(* IEC 61131-3 sources: codesys/project-view/Device/Plc Logic/Application/本机-3-机械臂-本体, 4 files *)

(* ---- Robot_STATE.st ---- *)
{attribute 'qualified_only'}
{attribute 'strict'}
(*A区三轴模组状态机*)
TYPE Robot_STATE :
(
	STOP := 0,						//停止
	INIT,						//初始化
	MANNUAL,					//手动模式
	AUTO,						//自动模式
	RobotAct,					//自动运行中
	MannualRun					//手动运行中
);
END_TYPE

(* ---- ST_ROBOT_MODULE.st ---- *)
TYPE ST_ROBOT_MODULE :	//机械臂模块
STRUCT
	bConnect					:BOOL;
	bConnected					:BOOL;
	bTcpError					:BOOL;

	//写
	x_iGrpEnable				:BOOL;			//上使能
	x_iGrpDisable				:BOOL;			//去使能
	x_iGrpReset					:BOOL;			//复位
	x_iStartScript				:BOOL;			//开始脚本
	x_iPauseScript				:BOOL;			//暂停脚本
	x_iContinueScript			:BOOL;			//继续脚本
	x_iStopScript				:BOOL;			//停止脚本
	x_iManualMode				:BOOL;			//手动模式
	x_iAutoMode					:BOOL;			//自动模式

	//读
	x_oStateRunning				:BOOL;			//状态-运行中
	x_oStateStopping			:BOOL;			//状态-停止中
	x_oStatePausing				:BOOL;			//状态-暂停中
	x_oStateFree				:BOOL;			//状态-空闲中
	x_oStateElectrify			:BOOL;			//状态-上电
	x_oStatePower				:BOOL;			//状态-使能中
	x_oStateErr					:BOOL;			//状态-报警
	x_oCollide					:BOOL;			//状态-碰撞

	//写
	wExecute_Init    			:WORD := 1;		//-- PLC请求初始化 (0/1)
	wExecute_Act     			:word;		//-- PLC请求执行动作 (0=无, 1=下料, 2=上料)
	wOrderNumCur     			:word;		//-- PLC指定工作站点 (1,2...)
	wRackTpye        			:word;		//-- PLC指定盘架类型
	wDeviceRackPosNum			:word;		//-- PLC指定设备取放编号
	wChassisRackPosNum			:WORD;		//-- PLC指定小车底盘位置编号
	xExcuteSetVal				:BOOL;		//搬运参数写入
	xExcuteInit					:BOOL;		//机械臂初始化
	xExcuteAct					:BOOL;		//执行机械臂搬运动作

	//读
	rGlobInitStatus				:WORD;			//初始化状态反馈		--4是初始化完成
	rOrderNumCur				:WORD;			//工作站点参数反馈
	rRackTpye					:WORD;			//盘架类型参数反馈
	rDeviceRackPosNum			:WORD;			//设备位置参数反馈
	rChassisRackPosNum			:WORD;			//小车位置参数反馈
	rAct_Status					:WORD;			//机械臂动作状态 (0=未执行,1=执行中,2=完成,3=失败)
	rExecute_Act				:WORD;			//当前执行动作反馈 (0=无, 1=下料, 2=上料)
	RobotBusy					:WORD;			//机械臂忙标志 (0=空闲, 1=忙碌)

	G_FailCode					:WORD;			//失败代码 (0=无错误, 1=RTU连接失败, 2=电爪初始化失败, 3=电爪打开失败, 4=电爪夹紧失败, 5=拍照失败)
	G_FailWorkstationrk			:WORD;			//失败时的工作站点编号
	G_FailActType				:WORD;			//失败时的动作类型 (1=下料/出库, 2=上料/入库)

END_STRUCT
END_TYPE

(* ---- Robot_ModbusClient.st ---- *)
PROGRAM Robot_ModbusClient
VAR_IN_OUT
	RobotMod							:ST_ROBOT_MODULE;
	Client								: ModbusFB.ClientTCP;
END_VAR
VAR_INPUT
	uiUnitId							: UINT:=1;		//设备ID
	udiTimeOut							: UDINT:=1000;	//动作时间，单位ms
	udiReplyTimeout						: UDINT:=1000;	//回复超时，单位ms
END_VAR
VAR

	FB_WriteSingleRegister				: ModbusFB.ClientRequestWriteSingleRegister;	//写单个寄存器 06
	FB_WriteMulRegister					: ModbusFB.ClientRequestWriteMultipleRegisters;	//写多个寄存器
	FB_ReadHoldingRegisters				: ModbusFB.ClientRequestReadHoldingRegisters;	//读保持寄存器 03
	FB_WriteSingleCoil 					: ModbusFB.ClientRequestWriteSingleCoil; 		//写单个线圈 05
	FB_ReadDiscreteInputs				: ModbusFB.ClientRequestReadDiscreteInputs;	//读触电寄存器  02
END_VAR
VAR
	Ton_LostConnect						: Standard.TON;
	bError								: BOOL;
	rTrig_Active						: Standard.R_TRIG;	//通讯连接成功上升沿
	iState								: INT;
END_VAR
VAR
	xDiscreteInputs						: ARRAY [0..11] OF BOOL;		//触电寄存器
	arrWHoldingRegisters				: ARRAY [0..7] OF WORD;
	arrWHoldingRegisters1				: ARRAY [0..2] OF WORD;
	arrWriteMulRegister					: ARRAY [0..3] OF WORD;

	pAction								:POINTER TO BOOL;
	Delay								:Standard.TON;
END_VAR
// --- implementation ---
ACT_01_FB();

ACT_02_Excute();

Act_03_State();

// (*断线、通讯错误时，自动重连*)
// IF ( NOT RobotMod.bConnected OR RobotMod.bTcpError OR bError ) AND RobotMod.bConnect THEN
// 	IF Ton_LostConnect.Q THEN
//         Ton_LostConnect(IN:=FALSE);
//     END_IF
//     Ton_LostConnect(IN:=TRUE, PT:=T#1000MS);
// ELSE
// 	Ton_LostConnect(IN:=FALSE);
// END_IF
END_PROGRAM

ACTION ACT_01_FB:
// Client(
// 	xConnected=> RobotMod.bTcpActive );

	(*客户端*)
//Client(xConnected=> RobotMod.bConnected);

//写单个寄存器
FB_WriteSingleRegister(
	xExecute:= ,
	udiTimeOut:= udiTimeOut * 1000, 				//单位us
	xDone=> ,
	xBusy=> ,
	xError=> ,
	rClient:= Client,
	uiUnitId:= uiUnitId,
	udiReplyTimeout:= udiReplyTimeout * 1000, 		//回复超时，单位us,
	uiMaxRetries:= ,
	eErrorID=> ,
	eException=> ,
	uiRetryCnt=> ,
	uiItem:= ,
	uiValue:= );

//写保持型寄存器
FB_ReadHoldingRegisters(
	xExecute:= ,
	udiTimeOut:= udiTimeOut * 1000, 				//单位us, ,
	xDone=> ,
	xBusy=> ,
	xError=> ,
	rClient:= Client,
	uiUnitId:= uiUnitId,
	udiReplyTimeout:= udiReplyTimeout * 1000, 		//回复超时，单位us, , ,
	uiMaxRetries:= ,
	eErrorID=> ,
	eException=> ,
	uiRetryCnt=> ,
	uiStartItem:= ,
	uiQuantity:= ,
	pData:= );

//写单个线圈
FB_WriteSingleCoil(
	xExecute:= ,
	udiTimeOut:= udiTimeOut * 1000, 				//单位us, ,
	xDone=> ,
	xBusy=> ,
	xError=> ,
	rClient:= Client,
	uiUnitId:= uiUnitId,
	udiReplyTimeout:= udiReplyTimeout * 1000, 		//回复超时，单位us, , ,
	uiMaxRetries:= ,
	eErrorID=> ,
	eException=> ,
	uiRetryCnt=> ,
	uiItem:= ,
	xValue:= );

//读取离散型输入
FB_ReadDiscreteInputs(
	xExecute:= ,
	udiTimeOut:= udiTimeOut * 1000, 				//单位us, ,
	xDone=> ,
	xBusy=> ,
	xError=> ,
	rClient:= Client,
	uiUnitId:= uiUnitId,
	udiReplyTimeout:= udiReplyTimeout * 1000, 		//回复超时，单位us, , ,
	uiMaxRetries:= ,
	eErrorID=> ,
	eException=> ,
	uiRetryCnt=> ,
	uiStartItem:= ,
	uiQuantity:= ,
	pData:= );

//写多个寄存器
FB_WriteMulRegister(
	xExecute:= ,
	udiTimeOut:=  udiTimeOut * 1000, 				//单位us, ,
	xDone=> ,
	xBusy=> ,
	xError=> ,
	rClient:= Client,
	uiUnitId:= uiUnitId,
	udiReplyTimeout:= udiReplyTimeout * 1000, 		//回复超时，单位us, , ,
	uiMaxRetries:= ,
	eErrorID=> ,
	eException=> ,
	uiRetryCnt=> ,
	uiStartItem:= ,
	uiQuantity:= , //“回复超时”情况下的请求重试次数。
	pData:= );
END_ACTION

ACTION ACT_02_Excute:
CASE iState OF
	0:
		//只读触点寄存器
		FB_ReadDiscreteInputs.uiStartItem := 0;
		FB_ReadDiscreteInputs.uiQuantity := 12;
		FB_ReadDiscreteInputs.pData := ADR(xDiscreteInputs);
		FB_ReadDiscreteInputs.xExecute := RobotMod.bConnected;
		IF FB_ReadDiscreteInputs.xDone THEN
			FB_ReadDiscreteInputs.xExecute:=FALSE;
			iState:=10;
		ELSIF FB_ReadDiscreteInputs.xError THEN
			iState:=1000;
		END_IF

	10:
		//读保持寄存器 1010-1017
		FB_ReadHoldingRegisters.uiStartItem := 1010;
		FB_ReadHoldingRegisters.uiQuantity := 8;
		FB_ReadHoldingRegisters.pData := ADR(arrWHoldingRegisters);
		FB_ReadHoldingRegisters.xExecute := RobotMod.bConnected;
		IF FB_ReadHoldingRegisters.xDone THEN
			FB_ReadHoldingRegisters.xExecute := FALSE;
			iState:=15;
		ELSIF FB_ReadHoldingRegisters.xError THEN
			iState:=1000;
		END_IF

	15:
		//读保持寄存器 1020-1022
		FB_ReadHoldingRegisters.uiStartItem := 1020;
		FB_ReadHoldingRegisters.uiQuantity := 3;
		FB_ReadHoldingRegisters.pData := ADR(arrWHoldingRegisters1);
		FB_ReadHoldingRegisters.xExecute := RobotMod.bConnected;
		IF FB_ReadHoldingRegisters.xDone THEN
			FB_ReadHoldingRegisters.xExecute := FALSE;
			iState:=20;
		ELSIF FB_ReadHoldingRegisters.xError THEN
			iState:=1000;
		END_IF

	20:
		//写运动指令
		//上使能
		IF RobotMod.x_iGrpEnable THEN
			pAction := ADR(RobotMod.x_iGrpEnable);
			FB_WriteSingleCoil.uiItem := 3;
			FB_WriteSingleCoil.xValue := TRUE;
			FB_WriteSingleCoil.xExecute := RobotMod.bConnected;
			IF FB_WriteSingleCoil.xDone THEN
				FB_WriteSingleCoil.xExecute := FALSE;
				iState:=50;
			ELSIF FB_WriteSingleCoil.xError THEN
				iState:=1000;
			END_IF
		//去使能
		ELSIF RobotMod.x_iGrpDisable THEN
			pAction := ADR(RobotMod.x_iGrpDisable);
			FB_WriteSingleCoil.uiItem := 4;
			FB_WriteSingleCoil.xValue := TRUE;
			FB_WriteSingleCoil.xExecute := RobotMod.bConnected;
			IF FB_WriteSingleCoil.xDone THEN
				FB_WriteSingleCoil.xExecute := FALSE;
				iState:=50;
			ELSIF FB_WriteSingleCoil.xError THEN
				iState:=1000;
			END_IF
		//清除报警
		ELSIF RobotMod.x_iGrpReset THEN
			pAction := ADR(RobotMod.x_iGrpReset);
			FB_WriteSingleCoil.uiItem := 5;
			FB_WriteSingleCoil.xValue := TRUE;
			FB_WriteSingleCoil.xExecute := RobotMod.bConnected;
			IF FB_WriteSingleCoil.xDone THEN
				FB_WriteSingleCoil.xExecute := FALSE;
				iState:=50;
			ELSIF FB_WriteSingleCoil.xError THEN
				iState:=1000;
			END_IF
		//开始脚本
		ELSIF RobotMod.x_iStartScript THEN
			pAction := ADR(RobotMod.x_iStartScript);
			FB_WriteSingleCoil.uiItem := 0;
			FB_WriteSingleCoil.xValue := TRUE;
			FB_WriteSingleCoil.xExecute := RobotMod.bConnected;
			IF FB_WriteSingleCoil.xDone THEN
				FB_WriteSingleCoil.xExecute := FALSE;
				iState:=50;
			ELSIF FB_WriteSingleRegister.xError THEN
				iState:=1000;
			END_IF
		//暂停脚本
		ELSIF RobotMod.x_iPauseScript THEN
			pAction := ADR(RobotMod.x_iPauseScript);
			FB_WriteSingleCoil.uiItem := 2;
			FB_WriteSingleCoil.xValue := TRUE;
			FB_WriteSingleCoil.xExecute := RobotMod.bConnected;
			IF FB_WriteSingleCoil.xDone THEN
				FB_WriteSingleCoil.xExecute := FALSE;
				iState:=50;
			ELSIF FB_WriteSingleCoil.xError THEN
				iState:=1000;
			END_IF
		//继续脚本
		ELSIF RobotMod.x_iContinueScript THEN
			pAction := ADR(RobotMod.x_iContinueScript);
			FB_WriteSingleCoil.uiItem := 2;
			FB_WriteSingleCoil.xValue := FALSE;
			FB_WriteSingleCoil.xExecute := RobotMod.bConnected;
			IF FB_WriteSingleCoil.xDone THEN
				FB_WriteSingleCoil.xExecute := FALSE;
				iState:=50;
			ELSIF FB_WriteSingleRegister.xError THEN
				iState:=1000;
			END_IF
		//停止脚本
		ELSIF RobotMod.x_iStopScript THEN
			pAction := ADR(RobotMod.x_iStopScript);
			FB_WriteSingleCoil.uiItem := 1;
			FB_WriteSingleCoil.xValue := TRUE;
			FB_WriteSingleCoil.xExecute := RobotMod.bConnected;
			IF FB_WriteSingleCoil.xDone THEN
				FB_WriteSingleCoil.xExecute := FALSE;
				iState:=50;
			ELSIF FB_WriteSingleCoil.xError THEN
				iState:=1000;
			END_IF
		//手动模式
		ELSIF RobotMod.x_iManualMode THEN
			pAction := ADR(RobotMod.x_iManualMode);
			FB_WriteSingleCoil.uiItem := 9;
			FB_WriteSingleCoil.xValue := TRUE;
			FB_WriteSingleCoil.xExecute := RobotMod.bConnected;
			IF FB_WriteSingleCoil.xDone THEN
				FB_WriteSingleCoil.xExecute := FALSE;
				iState:=50;
			ELSIF FB_WriteSingleCoil.xError THEN
				iState:=1000;
			END_IF
		//自动模式
		ELSIF RobotMod.x_iAutoMode THEN
			pAction := ADR(RobotMod.x_iAutoMode);
			FB_WriteSingleCoil.uiItem := 8;
			FB_WriteSingleCoil.xValue := TRUE;
			FB_WriteSingleCoil.xExecute := RobotMod.bConnected;
			IF FB_WriteSingleCoil.xDone THEN
				FB_WriteSingleCoil.xExecute := FALSE;
				iState:=50;
			ELSIF FB_WriteSingleCoil.xError THEN
				iState:=1000;
			END_IF
		//搬运参数写入	--iState 不需要跳 50
		ELSIF RobotMod.xExcuteSetVal THEN
			arrWriteMulRegister[0] 			:= RobotMod.wOrderNumCur;
			arrWriteMulRegister[1] 			:= RobotMod.wRackTpye;
			arrWriteMulRegister[2] 			:= RobotMod.wDeviceRackPosNum;
			arrWriteMulRegister[3] 			:= RobotMod.wChassisRackPosNum;
			FB_WriteMulRegister.uiStartItem := 1002;
			FB_WriteMulRegister.uiQuantity := 4;
			FB_WriteMulRegister.pData := ADR(arrWriteMulRegister);
			FB_WriteMulRegister.xExecute := RobotMod.bConnected;
			IF FB_WriteMulRegister.xDone THEN
				RobotMod.xExcuteSetVal := FALSE;
				FB_WriteMulRegister.xExecute := FALSE;
				iState:=100;
			ELSIF FB_WriteMulRegister.xError THEN
				iState:=1000;
			END_IF
		//执行初始化动作	--iState 不需要跳 50
		ELSIF RobotMod.xExcuteInit THEN
			FB_WriteSingleRegister.uiItem := 1000;
			FB_WriteSingleRegister.uiValue := 1;
			FB_WriteSingleRegister.xExecute := RobotMod.bConnected;
			IF FB_WriteSingleRegister.xDone THEN
				RobotMod.xExcuteInit := FALSE;
				FB_WriteSingleRegister.xExecute := FALSE;
				iState:=100;
			ELSIF FB_WriteSingleRegister.xError THEN
				iState:=1000;
			END_IF
		//执行搬运动作	--iState 不需要跳 50
		ELSIF RobotMod.xExcuteAct  THEN
			FB_WriteSingleRegister.uiItem := 1001;
			FB_WriteSingleRegister.uiValue := RobotMod.wExecute_Act;
			FB_WriteSingleRegister.xExecute := RobotMod.bConnected;
			IF FB_WriteSingleRegister.xDone THEN
				RobotMod.xExcuteAct := FALSE;
				FB_WriteSingleRegister.xExecute := FALSE;
				iState:=100;
			ELSIF FB_WriteSingleRegister.xError THEN
				iState:=1000;
			END_IF
		ELSE
			iState:=100;
		END_IF

		//线圈控制，仅上升沿有效，需要另外控制复位逻辑
	50:
		Delay(IN:= TRUE,PT:=T#50MS);
		IF Delay.Q THEN
			Delay(IN:= FALSE);
			FB_WriteSingleCoil.xValue := FALSE;
			FB_WriteSingleCoil.xExecute := RobotMod.bConnected;
			IF FB_WriteSingleCoil.xDone THEN
				FB_WriteSingleCoil.xExecute := FALSE;
				pAction^ := FALSE;
				iState:=100;
			ELSIF FB_WriteSingleCoil.xError THEN
				iState:=1000;
			END_IF
		END_IF

	100:
		bError:=FALSE;
		iState:=0;

	1000:
		bError := TRUE;
		FB_WriteSingleRegister.xExecute := FALSE;
		FB_WriteMulRegister.xExecute := FALSE;
		FB_ReadHoldingRegisters.xExecute := FALSE;
		FB_WriteSingleCoil.xExecute := FALSE;
		FB_ReadDiscreteInputs.xExecute := FALSE;

		Delay(IN:= TRUE,PT:=T#3S);
		IF Delay.Q THEN
			Delay(IN:= FALSE);
			iState:=0;
		END_IF
END_CASE
END_ACTION

ACTION Act_03_State:
RobotMod.x_oStateRunning :=xDiscreteInputs[0];
RobotMod.x_oStateStopping :=xDiscreteInputs[1];
RobotMod.x_oStatePausing :=xDiscreteInputs[2];
RobotMod.x_oStateFree :=xDiscreteInputs[5];
RobotMod.x_oStateElectrify := xDiscreteInputs[6];
RobotMod.x_oStatePower :=xDiscreteInputs[7];
RobotMod.x_oStateErr :=xDiscreteInputs[8];
RobotMod.x_oCollide :=xDiscreteInputs[9];

// -- 寄存器 1010-1017: 机械臂写入PLC的状态区域（机械臂写，PLC读）
// --   1010: GlobInitStatus   -- 初始化状态反馈
// --   1011: OrderNumCur      -- 当前工作站点反馈
// --   1012: RackTpye         -- 当前盘架类型反馈
// --   1013: DeviceRackPosNum -- 当前设备位置反馈
// --   1014: ChassisRackPosNum-- 当前小车位置反馈
// --   1015: Act_Status       -- 动作状态 (0=未执行,1=执行中,2=完成,3=失败)
// --   1016: Execute_Act      -- 当前执行动作反馈 (0/1/2)
// --   1017: RobotBusy        -- 机械臂忙标志 (0=空闲, 1=忙碌)
RobotMod.rGlobInitStatus 		:= arrWHoldingRegisters[0];
RobotMod.rOrderNumCur 			:= arrWHoldingRegisters[1];
RobotMod.rRackTpye	 			:= arrWHoldingRegisters[2];
RobotMod.rDeviceRackPosNum		:= arrWHoldingRegisters[3];
RobotMod.rChassisRackPosNum		:= arrWHoldingRegisters[4];
RobotMod.rAct_Status			:= arrWHoldingRegisters[5];
RobotMod.rExecute_Act			:= arrWHoldingRegisters[6];
RobotMod.RobotBusy				:= arrWHoldingRegisters[7];

// -- 寄存器 1020-1022: 失败详细信息（机械臂写，PLC读）
// --   1020: G_FailCode          -- 失败代码 (0=无错误, 1=RTU连接失败, 2=电爪初始化失败, 3=电爪打开失败, 4=电爪夹紧失败, 5=拍照失败)
// --   1021: G_FailWorkstationrk -- 失败时的工作站点编号
// --   1022: G_FailActType       -- 失败时的动作类型 (1=下料/出库, 2=上料/入库)
RobotMod.G_FailCode 			:= arrWHoldingRegisters[0];
RobotMod.G_FailWorkstationrk 	:= arrWHoldingRegisters[1];
RobotMod.G_FailActType 			:= arrWHoldingRegisters[2];
END_ACTION

(* ---- Robot_PRG.st ---- *)
PROGRAM Robot_PRG
VAR_IN_OUT
	Robot						: ST_ROBOT_MODULE;
END_VAR

VAR_INPUT
	bInitBtn					: BOOL;								//初始化按钮
	bStartBtn					: BOOL;								//启动按钮
	bPauseBtn					: BOOL;								//暂停按钮
	bStopBtn					: BOOL;								//停止按钮
	bResetBtn					: BOOL;								//复位按钮
	bAutoMode					: BOOL:= TRUE;						//true=自动模式，false=手动模式
END_VAR

VAR
	Warning_T					: Standard.TON;
	Warning						: BOOL;
	Delay						: Standard.TON;
END_VAR

//状态反馈
VAR

	wCommErrorCode				: WORD;	//通讯错误码
	wControllerState			: WORD;	//控制器状态机
	wInDriveSafe				: WORD;	//当前在行驶安全点(0:false，1:true)
	//wTaskID						: WORD;	//任务ID(当前任务ID，任务开始时获取一次，用于辨识)
	wTaskState					: WORD;	//任务状态(0:NONE，1:进行中，2:暂停中，3:已完成，4:参数异常，5:失败)
	wPhotoState					: WORD;	//拍照状态(0:空，1:拍照成功，2:拍照失败)
	wTakeRackState				: WORD;	//管架取料状态(0:空，1:抓料成功，2:抓料抓空，3:抓料抓歪)
	wPutRackState				: WORD;	//管架放料状态(0:空，1:放料成功，2:放料异常)
	wRackSensorState			: WORD;	//管架传感器状态(0:空，1:放料位被占用，2:取料位空闲)

	bMannualStart				: BOOL;		//手动模式启动

END_VAR

VAR
	eState						: Robot_STATE;						//总流程状态
	iInitStep					: INT;								//初始化步
	iAutoStep					: INT;								//自动步
	iMannualStep				: INT;								//手动模式步
	rTrig_Init					: Standard.R_TRIG;							//初始化按钮上升沿
	rTrig_Start					: Standard.R_TRIG;							//启动按钮上升沿
	rTrig_Pause					: Standard.R_TRIG;							//暂停按钮上升沿
	rTrig_Stop					: Standard.R_TRIG;							//停止按钮上升沿
	rTrig_Stop_1				: Standard.R_TRIG;							//停止按钮上升沿
	rTrig_Reset					: Standard.R_TRIG;							//复位按钮上升沿

END_VAR
VAR_OUTPUT
	iStepId						: INT;
	wsSteplog					: WSTRING;
	bBusy						: BOOL;								//正在运行标志位
	bInitializing				: BOOL;								//初始化中
	bInitialized				: BOOL;								//初始化完成标志位
	bAutoRunning				: BOOL;								//自动运行中
	bPausing					: BOOL;								//暂停中
	bStopping					: BOOL;								//停止中
	uliErrorId					: ULINT;							//错误ID
	uliWarningId				: ULINT;							//警告ID
	bReadyToRun					: BOOL;
	bOnSafePos					: BOOL;								//位于安全位置
END_VAR

VAR_INPUT

	uWorkStation				: UINT;		//工作站点
	uRackType					: UINT;		//管架类型
	uDeviceRackPos				: UINT;		//设备管架位置
	uChassisRackPos				: UINT;		//底盘管架位置
	wTaskID						: UINT;		//任务ID(ID标识符，用于辨识当前任务)
	wTaskNum					: UINT;		//工作方式 (0=无, 1=下料, 2=上料)
	bStart						: BOOL;
END_VAR
// --- implementation ---
bPausing := bPauseBtn;

ACT_00_FB();
Act_01_Stop();
ACT_02_State();
ACT_03_Warning();

(*初始化按钮*)
rTrig_Init(CLK:= bInitBtn);

CASE eState OF
	Robot_STATE.STOP:
		IF uliWarningId=0 AND uliErrorId=0  AND rTrig_Init.Q THEN		//停止模式下，进入初始化
		iInitStep := 0;
		bInitializing := TRUE;
		Act_99_ActionReset();
		eState := Robot_STATE.INIT;
	END_IF

	Robot_STATE.MANNUAL:
		bAutoRunning := FALSE;
		IF bMannualStart THEN
			eState := Robot_STATE.MannualRun;
		ELSIF bAutoMode THEN
			bAutoRunning := TRUE;
			eState := Robot_STATE.AUTO;
		END_IF

	Robot_STATE.INIT:
		Act_08_Init();
		IF bInitialized THEN		//初始化完成，进入自动模式
			bInitBtn := FALSE;
			bInitialized := FALSE;
			bAutoRunning := TRUE;
			eState := Robot_STATE.AUTO;
		END_IF

	Robot_STATE.MannualRun:
		ACT_11_bMannual();
		IF bAutoMode AND NOT bMannualStart AND iMannualStep = 0 THEN
			eState := Robot_STATE.AUTO;
		END_IF

	Robot_STATE.AUTO:
		IF uWorkStation>=1 AND uDeviceRackPos >= 1
			AND uChassisRackPos>=1 AND uChassisRackPos<=6 AND wTaskNum <> 0 AND bStart
				AND Glob_ModbusTcpServer.Car_xIsStatic
					AND NOT Glob_ModbusTcpServer.Car_xIsCharging
						AND NOT Glob_ModbusTcpServer.Car_xIsEStop THEN
			bBusy := TRUE;
			wTaskState := 1;
			iAutoStep := 0;
			eState := Robot_STATE.RobotAct;
		ELSIF NOT bAutoMode THEN
			eState := Robot_STATE.MANNUAL;
		END_IF

	Robot_STATE.RobotAct:
		ACT_10_RobotAct();
		IF NOT bBusy AND NOT bStart AND iAutoStep = 0 THEN
			eState := Robot_STATE.AUTO;
		END_IF

END_CASE
END_PROGRAM

ACTION Act_99_ActionReset:
iInitStep := 0;
iAutoStep := 0;
bBusy := FALSE;
bInitBtn := FALSE;
iMannualStep := 0;
END_ACTION

ACTION ACT_10_RobotAct:
CASE iAutoStep OF
	0:
		IF Robot.rGlobInitStatus = 4 AND Robot.rAct_Status <> 1 THEN
			Glob_ModbusTcpServer.Robot_wPhotoState := 0;
			iAutoStep := 10;
		END_IF

	10:
		//输入机器人参数
		Robot.wOrderNumCur := uWorkStation;
		Robot.wRackTpye := uRackType;
		Robot.wDeviceRackPosNum := uDeviceRackPos;
		Robot.wChassisRackPosNum := uChassisRackPos;
		Robot.xExcuteSetVal := TRUE;
		iAutoStep := 20;

	20:
		IF NOT Robot.xExcuteSetVal AND uWorkStation = Robot.rOrderNumCur
			AND uRackType = Robot.rRackTpye AND uDeviceRackPos = Robot.rDeviceRackPosNum
				AND uChassisRackPos = Robot.rChassisRackPosNum THEN
			iAutoStep := 30;
		END_IF

	30:
		//触发机器人动作
		Robot.wExecute_Act := wTaskNum;
		Robot.xExcuteAct := TRUE;
		iAutoStep := 40;

	40:
		IF NOT Robot.xExcuteAct AND  Robot.rAct_Status = 1 THEN
			iAutoStep := 50;
		END_IF

	50:
		//清空触发机器人动作
		Robot.wExecute_Act := 0;
		Robot.xExcuteAct := TRUE;
		iAutoStep := 60;

	60:
		IF NOT Robot.xExcuteAct THEN
			iAutoStep := 80;
		END_IF

		//机械臂状态写入
	80:
		IF Robot.rAct_Status = 2 AND NOT Robot.x_oStatePausing AND Robot.x_oStateRunning THEN	//运行完成
			Glob_ModbusTcpServer.Robot_wPhotoState := 1;
			Glob_ModbusTcpServer.Robot_wTaskState := 3;
			iAutoStep := 100;

		ELSIF Robot.rAct_Status = 3 OR uliWarningId <> 0 THEN	//报错
			//Glob_ModbusTcpServer.Robot_wTaskState := 5;
			iAutoStep := 85;

		ELSIF Robot.rAct_Status = 1 AND NOT Robot.x_oStatePausing THEN
			Glob_ModbusTcpServer.Robot_wTaskState := 1;

		ELSIF Robot.rAct_Status = 1 AND Robot.x_oStatePausing THEN
			Glob_ModbusTcpServer.Robot_wTaskState := 2;

		END_IF

	85:
		Glob_ModbusTcpServer.Robot_wTaskState := 5;
		IF Robot.G_FailCode = 5 THEN
			Glob_ModbusTcpServer.Robot_wPhotoState := 2;
		END_IF
		iAutoStep := 100;

	100:
		//清空触发机器人动作
		Robot.wExecute_Act := 0;
		Robot.xExcuteAct := TRUE;
		iAutoStep := 150;

	150:
		IF NOT Robot.xExcuteAct AND  Robot.rAct_Status <> 1 THEN
			iAutoStep := 500;
		END_IF

	500:
		wTaskNum := 0;
		uWorkStation := 0;
		uRackType := 0;
		uDeviceRackPos := 0;
		uChassisRackPos := 0;
		bStart := FALSE;
		bBusy := FALSE;
		iAutoStep := 0;
END_CASE
END_ACTION

ACTION ACT_00_FB:
END_ACTION

ACTION Act_01_Stop:
(*停止按钮*)
rTrig_Stop(CLK :=  bStopBtn);
IF rTrig_Stop.Q THEN
	eState := Robot_STATE.STOP;
END_IF

(*停止状态标志位*)
IF eState=Robot_STATE.STOP THEN

	bInitializing := FALSE;
	bInitialized := FALSE;
	bAutoRunning := FALSE;
	bPausing := FALSE;
	bStopping := TRUE;
	Delay(IN:= FALSE);
	iAutoStep := 0;
	bStart := FALSE;
	bBusy := FALSE;
	iStepId := 2;

	wsSteplog := "急停中，等待复位初始化";
ELSE
	bStopping := FALSE;
END_IF

rTrig_Stop_1(CLK :=  eState=Robot_STATE.STOP);
IF rTrig_Stop_1.Q THEN
	Robot.x_iStopScript := TRUE;
	Robot.x_iGrpDisable := TRUE;
END_IF
END_ACTION

ACTION Act_08_Init:
CASE iInitStep OF
	0:
		Robot.bConnect := TRUE;
		Glob.Chassis_Car.bConnect := TRUE;
		Robot.x_iAutoMode := FALSE;
		Warning_T(IN := TRUE,PT:= T#5S);
		IF Robot.bConnected AND Glob.Chassis_Car.bConnected THEN
			Warning_T(IN := FALSE);
			iInitStep := 20;
		ELSIF Warning_T.Q THEN
			;
		END_IF

		//机械臂切换手动模式
	20:
		Robot.x_iAutoMode := TRUE;
		Delay(IN := TRUE,PT := T#500MS);
		IF Delay.Q THEN
			Delay(IN := false);
			iInitStep := 30;
		END_IF

	30:
		IF NOT Robot.x_iAutoMode THEN
			iInitStep := 50;
		END_IF

		//机械臂运行脚本
	50:
		IF NOT Robot.x_oStatePower THEN
			Robot.x_iGrpEnable := TRUE;
		ELSIF Robot.x_oStateErr THEN
			Robot.x_iGrpReset := TRUE;
		ELSIF Robot.x_oStateFree OR Robot.x_oStateStopping THEN
			Robot.x_iStartScript := TRUE;
		ELSIF Robot.x_oStatePausing THEN
			Robot.x_iStopScript := TRUE;
		ELSIF Robot.x_oStateRunning THEN
			iInitStep := 100;
		END_IF

	100:
		Delay(IN := TRUE,PT := T#1000MS);
		IF Delay.Q THEN
			Delay(IN := false);
			iInitStep := 105;
		END_IF

	105:
		//机械臂运行初始化动作
		//Robot.wExecute_Init := 1;
		Robot.xExcuteInit := TRUE;
		Delay(IN := TRUE,PT := T#1000MS);
		IF Delay.Q THEN
			Delay(IN := false);
			iInitStep := 110;
		END_IF

	110:
		IF NOT Robot.xExcuteInit THEN
			iInitStep := 120;
		END_IF

	120:
		IF Robot.rGlobInitStatus = 4 THEN
			iInitStep := 150;
		END_IF

	150:
		Robot.wExecute_Act := 0;
		Robot.xExcuteAct := TRUE;
		iInitStep := 160;

	160:
		IF NOT Robot.xExcuteAct AND  Robot.rAct_Status = 0 THEN
			iInitStep := 1000;
		END_IF

	1000:
		iStepId := 1;
		wsSteplog := "待机中";

		bInitializing := FALSE;
		bInitialized := TRUE;
		iInitStep := 0;

END_CASE
END_ACTION

ACTION ACT_02_State:
END_ACTION

ACTION ACT_03_Warning:
IF eState = Robot_STATE.AUTO OR eState = Robot_STATE.RobotAct THEN

	uliWarningId.1 S= NOT Robot.bConnected;				//机械臂TCP未连接
	uliWarningId.2 S= Robot.bTcpError;					//机械臂TCP功能块错误
	uliWarningId.3 S= Robot.x_oStateErr;				//机械臂-报警
	uliWarningId.4 S= Robot.x_oCollide;					//机械臂-碰撞
	uliWarningId.5 S= Robot.x_oStateStopping;			//机械臂-停止运行
	uliWarningId.6 S= NOT Robot.x_oStateElectrify;		//机械臂-未上电
	uliWarningId.7 S= NOT Robot.x_oStatePower;			//机械臂-未使能
	uliWarningId.8 S= NOT Robot.x_oStateRunning;		//未运行
	uliWarningId.9 S= Robot.rGlobInitStatus <> 4;		//未初始化

	IF uliWarningId<>0 AND eState = Robot_STATE.RobotAct THEN
		Glob_ModbusTcpServer.Robot_wTaskState := 5;
		eState := Robot_STATE.STOP;
	ELSIF uliWarningId<>0 AND eState = Robot_STATE.AUTO THEN
		eState := Robot_STATE.STOP;
	END_IF

END_IF

(*复位按钮*)
rTrig_Reset(CLK :=  bResetBtn);
IF rTrig_Reset.Q THEN
	uliWarningId := 0;
END_IF
END_ACTION

ACTION ACT_11_bMannual:
CASE iMannualStep OF
	0:
		IF bMannualStart THEN
			iMannualStep := 10;
		END_IF

	10:
		Robot.xExcuteAct := TRUE;
		iMannualStep := 20;

	20:
		IF NOT Robot.xExcuteAct AND  Robot.rAct_Status = 1 THEN
			iMannualStep := 50;
		END_IF

	50:
		//清空触发机器人动作
		Robot.wExecute_Act := 0;
		Robot.xExcuteAct := TRUE;
		iMannualStep := 60;

	60:
		IF NOT Robot.xExcuteAct THEN
			iMannualStep := 1000;
		END_IF

	1000:
		bMannualStart := FALSE;
		iMannualStep := 0;
END_CASE
END_ACTION
